(* IEC 61131-3 sources: SortJet_MasterSPS_Aufbau.fbsproj/Device.device.xml.v3^/Plc Logic.plclogic.xml.v3^/Application.application.xml.v3^/09_Station/Shuttle/[151,152] Transfershuttle/0_Konfig, 6 files *)

(* ---- Antriebsinformationen_151.gvl ---- *)
(* METADATA
{
	"v3Meta": {
		"objectGuid": "1be33521-6e58-4da8-829e-a9c5887a7afb"
	}
}
*)
{attribute 'allow_unqualified_access'}
NAMESPACE Antriebsinformationen_151
VAR_GLOBAL

//-------------------------------------------------------------------------------------------------
// ANTRIEBSINFORMATION TRANSFERSHUTTLE
//-------------------------------------------------------------------------------------------------

  apgInfoTransfershuttle151Querfahrt : AntriebsInformationen :=
    (
      wAchsID                                 :=         0,  // Achs ID aus dem EConSet
      stTyp                                   := 'Lateral',  // Typ
      wpSchaltschrank                         :=         2,  // Daten aus dem Schaltplan
      wpSchaltplanreihe                       :=         2,  // Daten aus dem Schaltplan
      wpSchaltplanseite                       :=        60,  // Daten aus dem Schaltplan
      rpMaxGeschwindigkeit                    :=      3333,  // [mm/s]   Max- Geschwindigkeit für den Automatikbetrieb
      rpHandGeschwindigkeit                   :=       200,  // [mm/s]   Hand- Geschwindigkeit
      rpReferenzGeschwindigkeit               :=        50,  // [mm/s]   Geschwindigkeit für die Referenzfahrt
      rpMaxBeschleunigung                     :=      4000,  // [mm/s^2] Max Beschleunigung
      rpMaxVerzoegerung                       :=      4000,  // [mm/s^2] Max Verzoegerung
      rpMaxRuckzeit                           :=       300,  // [ms]     Ruckzeit des Antriebs
      rpReduzierteBeschleunigung              :=      4000,  // [mm/s^2] Reduzierte Beschleunigung
      rpReduzierteVerzoegerung                :=      4000,  // [mm/s^2] Reduzierte Verzoegerung
      rpEinrichtGeschwindigkeit               :=        50,  // [mm/s]   Max Geschwindigkeit während der Einrichtung der Anlage
      rpReduzierteGeschwindigkeit             :=       0.0,  // [mm/s]   Reduzierte Geschwindigkeit
      rpBeschleunigungFremdanlage             :=       0.0,  // [mm/s^2] Beschleunigung zu einer Fremdanlage
      rpGeschwindigkeitMessen                 :=       0.0,  // [mm/s] Geschwindigkeit beim Scheiben messen
      rpGeschwindigkeitSystemcheck            :=     500.0,  // [mm/s]   Geschwindigkeit im Systemcheck (nur Glastransport)
      rpGeschwindigkeitSystemcheckReduzierung :=     167.0,  // [mm/s]   Geschwindigkeit im Systemcheck bei belegtem Vorstop-Sensor (nur Glastransport)
      stOptionen                              := ( eEndschalterQuelle    := Endschalterquelle_EN.UMRICHTER, // Hardware-Endschalter: KEINE, UMRICHTER oder SPS
                                                   bVersorgungUeberXVR   := FALSE,                          // XVR-Modus: brueckt Hauptschalter 400 V und LS 230 V
                                                   bBremseLoesenFreigabe := FALSE )                         // Der Antrieb darf über eine Betriebsart die Bremse lösen
    );

  apgInfoTransfer151Glastransport : ARRAY[cWAND_1..cANZAHL_WAENDE] OF AntriebsInformationen := [
    (
      wAchsID                                 :=         1,  // Achs ID aus dem EConSet
      stTyp                                   :=    'Belt',  // Typ
      wpSchaltschrank                         :=         2,  // Daten aus dem Schaltplan
      wpSchaltplanreihe                       :=         2,  // Daten aus dem Schaltplan
      wpSchaltplanseite                       :=        65,  // Daten aus dem Schaltplan
      rpMaxGeschwindigkeit                    :=       667,  // [mm/s]   Max- Geschwindigkeit für den Automatikbetrieb
      rpHandGeschwindigkeit                   :=       200,  // [mm/s]   Hand- Geschwindigkeit
      rpReduzierteGeschwindigkeit             :=        67,  // [mm/s]   Reduzierte Geschwindigkeit
      rpReferenzGeschwindigkeit               :=         0,  // [mm/s]   Geschwindigkeit für die Referenzfahrt
      rpEinrichtGeschwindigkeit               :=        50,  // [mm/s]   Max Geschwindigkeit während der Einrichtung der Anlage
      rpMaxBeschleunigung                     :=      1500,  // [mm/s^2] Max Beschleunigung
      rpMaxVerzoegerung                       :=      2000,  // [mm/s^2] Max Verzoegerung
      rpMaxRuckzeit                           :=        50,  // [ms]     Ruckzeit des Antriebs
      rpReduzierteBeschleunigung              :=      1000,  // [mm/s^2] Reduzierte Beschleunigung
      rpReduzierteVerzoegerung                :=      1000,  // [mm/s^2] Reduzierte Verzoegerung
      rpBeschleunigungFremdanlage             :=      1000,  // [mm/s^2] Beschleunigung zu einer Fremdanlage
      rpGeschwindigkeitMessen                 :=       667,  // [mm/s] Geschwindigkeit beim Scheiben messen
      rpGeschwindigkeitSystemcheck            :=     500.0,  // [mm/s]   Geschwindigkeit im Systemcheck (nur Glastransport)
      rpGeschwindigkeitSystemcheckReduzierung :=     167.0,  // [mm/s]   Geschwindigkeit im Systemcheck bei belegtem Vorstop-Sensor (nur Glastransport)
      stOptionen                              := ( eEndschalterQuelle    := Endschalterquelle_EN.KEINE,     // Hardware-Endschalter: KEINE, UMRICHTER oder SPS
                                                   bVersorgungUeberXVR   := FALSE,                          // XVR-Modus: brueckt Hauptschalter 400 V und LS 230 V
                                                   bBremseLoesenFreigabe := FALSE )                         // Der Antrieb darf über eine Betriebsart die Bremse lösen
    )];

END_VAR
END_NAMESPACE

(* ---- Antriebsinformationen_152.gvl ---- *)
(* METADATA
{
	"v3Meta": {
		"objectGuid": "34921d73-d8bd-4657-bcb2-03b0c8f4301f"
	}
}
*)
{attribute 'allow_unqualified_access'}
NAMESPACE Antriebsinformationen_152
VAR_GLOBAL

//-------------------------------------------------------------------------------------------------
// ANTRIEBSINFORMATION TRANSFERSHUTTLE
//-------------------------------------------------------------------------------------------------

  apgInfoTransfershuttle152Querfahrt : AntriebsInformationen :=
    (
      wAchsID                                 :=         2,  // Achs ID aus dem EConSet
      stTyp                                   := 'Lateral',  // Typ
      wpSchaltschrank                         :=         2,  // Daten aus dem Schaltplan
      wpSchaltplanreihe                       :=         2,  // Daten aus dem Schaltplan
      wpSchaltplanseite                       :=        60,  // Daten aus dem Schaltplan
      rpMaxGeschwindigkeit                    :=      3333,  // [mm/s]   Max- Geschwindigkeit für den Automatikbetrieb
      rpHandGeschwindigkeit                   :=       200,  // [mm/s]   Hand- Geschwindigkeit
      rpReferenzGeschwindigkeit               :=        50,  // [mm/s]   Geschwindigkeit für die Referenzfahrt
      rpMaxBeschleunigung                     :=      4000,  // [mm/s^2] Max Beschleunigung
      rpMaxVerzoegerung                       :=      4000,  // [mm/s^2] Max Verzoegerung
      rpMaxRuckzeit                           :=       300,  // [ms]     Ruckzeit des Antriebs
      rpReduzierteBeschleunigung              :=      4000,  // [mm/s^2] Reduzierte Beschleunigung
      rpReduzierteVerzoegerung                :=      4000,  // [mm/s^2] Reduzierte Verzoegerung
      rpEinrichtGeschwindigkeit               :=        50,  // [mm/s]   Max Geschwindigkeit während der Einrichtung der Anlage
      rpReduzierteGeschwindigkeit             :=       0.0,  // [mm/s]   Reduzierte Geschwindigkeit
      rpBeschleunigungFremdanlage             :=       0.0,  // [mm/s^2] Beschleunigung zu einer Fremdanlage
      rpGeschwindigkeitMessen                 :=       0.0,  // [mm/s] Geschwindigkeit beim Scheiben messen
      rpGeschwindigkeitSystemcheck            :=     500.0,  // [mm/s]   Geschwindigkeit im Systemcheck (nur Glastransport)
      rpGeschwindigkeitSystemcheckReduzierung :=     167.0,  // [mm/s]   Geschwindigkeit im Systemcheck bei belegtem Vorstop-Sensor (nur Glastransport)
      stOptionen                              := ( eEndschalterQuelle    := Endschalterquelle_EN.UMRICHTER, // Hardware-Endschalter: KEINE, UMRICHTER oder SPS
                                                   bVersorgungUeberXVR   := FALSE,                          // XVR-Modus: brueckt Hauptschalter 400 V und LS 230 V
                                                   bBremseLoesenFreigabe := FALSE )                         // Der Antrieb darf über eine Betriebsart die Bremse lösen
    );

  apgInfoTransfer152Glastransport : ARRAY[cWAND_1..cANZAHL_WAENDE] OF AntriebsInformationen := [
    (
      wAchsID                                 :=         3,  // Achs ID aus dem EConSet
      stTyp                                   :=    'Belt',  // Typ
      wpSchaltschrank                         :=         2,  // Daten aus dem Schaltplan
      wpSchaltplanreihe                       :=         2,  // Daten aus dem Schaltplan
      wpSchaltplanseite                       :=        65,  // Daten aus dem Schaltplan
      rpMaxGeschwindigkeit                    :=       667,  // [mm/s]   Max- Geschwindigkeit für den Automatikbetrieb
      rpHandGeschwindigkeit                   :=       200,  // [mm/s]   Hand- Geschwindigkeit
      rpReduzierteGeschwindigkeit             :=        67,  // [mm/s]   Reduzierte Geschwindigkeit
      rpReferenzGeschwindigkeit               :=         0,  // [mm/s]   Geschwindigkeit für die Referenzfahrt
      rpEinrichtGeschwindigkeit               :=        50,  // [mm/s]   Max Geschwindigkeit während der Einrichtung der Anlage
      rpMaxBeschleunigung                     :=      1500,  // [mm/s^2] Max Beschleunigung
      rpMaxVerzoegerung                       :=      2000,  // [mm/s^2] Max Verzoegerung
      rpMaxRuckzeit                           :=        50,  // [ms]     Ruckzeit des Antriebs
      rpReduzierteBeschleunigung              :=      1000,  // [mm/s^2] Reduzierte Beschleunigung
      rpReduzierteVerzoegerung                :=      1000,  // [mm/s^2] Reduzierte Verzoegerung
      rpBeschleunigungFremdanlage             :=      1000,  // [mm/s^2] Beschleunigung zu einer Fremdanlage
      rpGeschwindigkeitMessen                 :=       667,  // [mm/s] Geschwindigkeit beim Scheiben messen
      rpGeschwindigkeitSystemcheck            :=     500.0,  // [mm/s]   Geschwindigkeit im Systemcheck (nur Glastransport)
      rpGeschwindigkeitSystemcheckReduzierung :=     167.0,  // [mm/s]   Geschwindigkeit im Systemcheck bei belegtem Vorstop-Sensor (nur Glastransport)
      stOptionen                              := ( eEndschalterQuelle    := Endschalterquelle_EN.KEINE,     // Hardware-Endschalter: KEINE, UMRICHTER oder SPS
                                                   bVersorgungUeberXVR   := FALSE,                          // XVR-Modus: brueckt Hauptschalter 400 V und LS 230 V
                                                   bBremseLoesenFreigabe := FALSE )                         // Der Antrieb darf über eine Betriebsart die Bremse lösen
    )];

END_VAR
END_NAMESPACE

(* ---- MK_Transfershuttle_151.gvl ---- *)
(* METADATA
{
	"v3Meta": {
		"objectGuid": "7b0b09af-66f3-4d35-ae87-7c9d4c69f207"
	}
}
*)
{attribute 'allow_unqualified_access'}
NAMESPACE MK_Transfershuttle_151
VAR_GLOBAL

//-------------------------------------------------------------------------------------------------
// TRANSFERSHUTTLE ALLGEMEIN
//-------------------------------------------------------------------------------------------------

  apgMKTransfershuttle151 : Parameter_Station :=
    (
      stStationsNummern                 := ( NummerIntern := 151,                                     // Stationsnummer fuer das MMI und die Stationsangabe der Meldungen
                                             NummerExtern := 1151,                                    // Stationsnummer fuer Bedienermeldungen
                                             NummerSPS    := 151 ),                                   // Stationsnummer SPS-intern (Indizes)
      bDeaktivieren                     := FALSE,                                                     // Station deaktiviert (keine Auftraege, keine Referenzfahrt)
      wMeldungsNummer                   := 350,                                                       // Basis-Meldungsnummer (WatchIO)
      eStationsTyp                      := eTransfershuttle,                                          // Typ der Station
      eaAutomatikkreis                  := [eAutomatikkreis_1, eAutomatikkreis_2],                    // Automatikkreise, zu denen die Station gehoert
      eaSicherheitskreis                := [eSicherheitskreis_1],                                     // Sicherheitskreise, in die die Station eingebunden ist
      // astSicherheitskreisTeilabschaltung
      eSystemcheckZyklus                := eSystemcheckZyklus_1,                                      // In welchem Zyklus des Systemchecks die Station geprueft wird
      stSchnittstellendaten             := ( wVorgaengerStation := cSTATION_DEFAULT,                  // Station vor dieser Station (cSTATION_DYNAMISCH bei mehreren)
                                             wNachfolgerStation := cSTATION_DEFAULT,                  // Station nach dieser Station (cSTATION_DYNAMISCH bei mehreren)
                                             bStationIstShuttle := TRUE ),                            // Station ist ein Shuttle

      stStationsOptionen                := (
                                            stSystemcheck := (
                                              bScheibenVermessenSystemCheck           := FALSE,       // Scheiben im Systemcheck vermessen
                                              bScheibeNachSystemcheckAufAuslauf       := FALSE,       // Scheibe nach dem Systemcheck auf den Auslaufsensor fahren
                                              bSystemCheckMitVorgaengerBatchTransport := FALSE,       // derzeit ohne Funktion
                                              bSystemCheckMitNachfolgerBatchTransport := FALSE,       // derzeit ohne Funktion
                                              bOptionSystemCheckScheibeMittigLegen    := FALSE        // derzeit ohne Funktion
                                            ),

                                            stTransfershuttle := (
                                              bMasterStation                          := TRUE,        // Ob es sich um ein Master (Master-Slave) - Station handelt. Aktuell gebraucht bei Transfershuttle- Verbund
                                              bTransferShuttleFuerFaecherwagen        := FALSE,       // Transfershuttle beschickt Faecherwagen
                                              bTransferShuttleMitUltraschallSensoren  := FALSE,       // Luftabfragen als Ultraschallsensoren (Schliesser)
                                              bTransfershuttleIstVerfahrbarerSpeicher := FALSE        // Transfershuttle ist verfahrbarer Speicher
                                            ),

                                            stGlastransport := (
                                              bVortransport                          := TRUE,         // Vortransport aktivieren [Bsp.: Nach einem Eintransport mit gesetztem Bit <Letzte Scheibe>]
                                              bTransportMasterSlaveEintransport      := FALSE,        // derzeit ohne Funktion
                                              bTransportMasterSlaveAustransport      := TRUE ,        // Austransport als Slave auf die Achse des Nachfolgers
                                              bGLasUebernahmeSenkrecht               := FALSE,        // RKT - Eintransport in Senkrechter-Position bzw. in Waagerechter- Position [default]
                                              bAustransportISOLinie                  := FALSE,        // Austransport an eine ISO-Linie
                                              bScheibenVermessen                     := FALSE,        // Scheibenmessung am Anlegetisch/Anlegewand
                                              bMessrichtungNegativ                   := FALSE,        // Negative Fahrtrichtung beim Messen
                                              bScheibenmessungEintransport           := FALSE,        // Scheibenmessung beim Eintransport
                                              bScheibenmessungSensorVorabAuslauf     := FALSE         // Scheibenmessung mit SensorVorabAuslauf z.B. Anlegewand
                                            ),

                                            // stAnlegetisch
                                            // stEckuebergabe
                                            // stDrehstation
                                            bVorAbKomponentenAnsteuerung            := FALSE,         // VorAbKomponentenAnsteuerung Auftraege werden bearbeitet
                                            bVerstellungEinAusGefahrenLogikDrehen   := FALSE,         // Verstellung: Logik ein-/ausgefahren gedreht
                                            bLangsamfahrtNockenQuerfahrtAktivieren  := FALSE,         // Querfahrt: Langsamfahrt-Nocken auswerten
                                            bSKBlockierenDurchVorabSensoren         := FALSE,         // Vorab-Sensoren belegt blockieren das Oeffnen des Sicherheitskreises
                                            bStationLeerfahrenBeiSkAnforderung      := FALSE,         // Station bei Anforderung Sicherheitskreis leerfahren
                                            bGlasAbgenommenAutomatischQuittieren    := FALSE,         // derzeit ohne Funktion
                                            bScheibeAbnehmenNachEintransport        := FALSE          // Scheibe nach dem Eintransport wieder abnehmen
                                          ),

      stStationsAufbau                  := (
                                            bGeblase                      := [cANZAHL_WAENDE(FALSE)], // Ausbaustufe: Geblaese je Wand
                                            bGlastransport                := [cANZAHL_WAENDE(TRUE)],  // Ausbaustufe: Glastransport je Wand
                                            bKippen                       := [cANZAHL_WAENDE(FALSE)], // Ausbaustufe: Kippen je Wand
                                            bKippenSchuetz                := FALSE,                   // Kippen ueber Schuetz statt Umrichter
                                            bTransportVerstellung         := [cANZAHL_WAENDE(FALSE)], // Ausbaustufe Shuttle: Transport-/Dickenverstellung je Wand
                                            bHub                          := FALSE,                   // Ausbaustufe: Hub der Station
                                            bHubrahmen                    := FALSE,                   // Ausbaustufe: Hubrahmen (Riemen heben/senken)
                                            bDrehen                       := FALSE,                   // Ausbaustufe: Drehen
                                            bQuerachse                    := FALSE,                   // Ausbaustufe: Querachse
                                            bMessachse                    := FALSE,                   // Ausbaustufe: Messachse (Anlegetisch, Anlegewand)
                                            bDruckluft                    := TRUE,                    // Druckluftueberwachung vorhanden
                                            bAnschlag                     := FALSE,                   // Ausbaustufe: Ausrichtanschlaege
                                            bSensorAuslauf                := TRUE,                    // Auslaufsensor vorhanden
                                            bSensorEinlauf                := TRUE,                    // Einlaufsensor vorhanden
                                            bSensorEinlaufStopp           := FALSE,                   // Shuttle: zusaetzlicher Stopp-Sensor am Einlauf (ohne: Einlaufsensor), Gegenstueck zum Auslauf-Stopp im Rueckwaertstransport
                                            bSensorAuslaufStopp           := FALSE,                   // Shuttle: zusaetzlicher Stopp-Sensor am Auslauf (ohne: Auslaufsensor), Verfahrfreigabe und Scheibe hat Shuttle verlassen
                                            bDurchlaufSperreZumNachfolger := FALSE,                   // Ausbaustufe: bewegliche Abschrankung zum Nachfolger
                                            bQuerfahrt                    := TRUE,                    // Ausbaustufe: Querfahrt
                                            bDLSSchmiersystem             := TRUE,                    // Zentralschmierung DLS vorhanden
                                            bWandverstellung              := [ FALSE ],               // Ausbaustufe Station: Wandverstellung je Wand
                                            bWandverstellungMotorisch     := FALSE,                   // Shuttle: Transport-/Wandverstellung mit Antrieb statt pneumatisch
                                            bRoellchenleiste              := [ FALSE ],               // Ausbaustufe Station: Roellchenleiste je Wand
                                            bDurchgang                    := FALSE,                   // Station ist Teil eines Durchgangs (belegt = Oeffnen blockiert)
                                            bSlaveAntrieb                 := FALSE,                   // Glastransport mit Slave-Antrieb
                                            bRolltor                      := FALSE,                   // Ausbaustufe Faecherwagen: Rolltor
                                            bKlemmzylinder                := FALSE,                   // Ausbaustufe Faecherwagen: Klemmzylinder fixiert den Oberrahmen beim Ein- und Ausschleusen
                                            bGreifer                      := [cANZAHL_WAENDE(FALSE)], // Shuttle: Greifer je Wand (Scheibe aus dem Faecherwagen ziehen bzw. hineinschieben)
                                            bRFID                         := FALSE,                   // RFID-Leser vorhanden
                                            bAGV                          := FALSE,                   // Ausbaustufe Faecherwagen: Betrieb mit AGV
                                            bKipparme                     := FALSE,                   // Ausbaustufe: Kipparme
                                            bMessachseAmEndeVomTisch      := FALSE,                   // Messachse am Ende des Tisches (Hoehenfehler fragt den Bediener)
                                            bGlastransportSlaveVorhanden  := FALSE,                   // Glastransport mit Slave-Antrieb (Meldungen/Ueberwachung Slave)
                                            wHydraulikstation             := 0                        // Faecherwagen Hydraulik: zugeordnete Hydraulikstation (cHYDRAULIKSTATION_x), 0 = keine
                                          ),

      stStationsParameter               := (
                                            rLaengeUebergroesseScheibe              := 4240,          // Shuttle: ab dieser Scheibenlaenge gilt die Scheibe als uebergross [mm]
                                            rMinGlasHoeheAutomatischenEintransport  := 500,           // VSG: Mindesthoehe fuer automatischen Eintransport [mm]
                                            rMinGlasLaengeAutomatischenEintransport := 500,           // VSG: Mindestlaenge fuer automatischen Eintransport [mm]
                                            wMaximaleAnzahlAktiverAuftraege         := 1,             // derzeit ohne Funktion
                                            rMinPosSwEsEingrenzung                  := 0.0,           // Externer zusaetzlicher Software-Endschalter MIN; 0 = inaktiv; darf den MK-MIN nur weiter eingrenzen
                                            rMaxPosSwEsEingrenzung                  := 0.0,           // Externer zusaetzlicher Software-Endschalter MAX; 0 = inaktiv; darf den MK-MAX nur weiter eingrenzen
                                            rPosFreigabePufferAusfahren             := 0.0            // derzeit ohne Funktion
                                          ),

      // stFremdanlage
      stGlasdaten                       := [
                                            (
                                              rlMinGlasLaenge := 350,                                 // minimal zulässige GlasLänge
                                              rlMaxGlasLaenge := 2500,                                // maximale zulässige GlasLänge
                                              rlMinGlasHoehe  := 190,                                 // minimal zulässige GlasHöhe
                                              rlMaxGlasHoehe  := 1800,                                // maximale zulässige GlasHöhe
                                              rlMinGlasDicke  := 3,                                 // minimal zulässige GlasDicke
                                              rlMaxGlasDicke  := 12.76,                                  // maximal zulaessige Glasdicke [mm]
                                              rlLaengeMaxGlas := 0.0                                  // maximal zulaessige Glaslaenge [mm]
                                            )]
      // astShuttleAnhaltenQuellen
    );

//-------------------------------------------------------------------------------------------------
// TRANSFERSHUTTLE GLASTRANSPORT
//-------------------------------------------------------------------------------------------------

  apgTransfer151Glastransport : ARRAY[cWAND_1..cANZAHL_WAENDE] OF Parameter_TransfershuttleGlastransport := [
    (
      rlLaengeStation                    := 3945, // Länge der Station
      rStopFreiFahren                    := 300,  // So weit soll die Scheibe beim Austransport länger fahren
      rWegUeberEinlaufEintransport       := 170,  // Eintransport vorwaerts: Abstand Scheibenhinterkante zum Einlaufsensor [mm]
      rWegUeberEinlaufAustransport       := 50,   // Lage Auf Einlauf: Scheibe liegt um diesen Weg auf dem Einlaufsensor [mm]
      rWegUeberAuslaufEintransport       := 50,   // Eintransport rueckwaerts: Abstand Scheibenhinterkante zum Auslaufsensor [mm]
      rWegUeberAuslaufAustransport       := 50,   // Lage Auf Auslauf: Weg ueber den Auslaufsensor hinaus [mm]
      wEnergieSparZeit                   := 180,  // in Sec, Zeitspanne nach der, der Antrieb deaktiviert wird wenn er keinen Auftrag hat
      rMaxPosAuslaufSensorFreiFahren     := 300,  // Bestimmt die Strecke die Maximal zurueck gefahren werden soll bis der Auslaufsensor  wieder frei ist
      rMaxPosEinlaufSensorFreiFahren     := 300,  // So weit darf maximal der Einlaufsensor frei gefahren weirden
      rgAbstandLuftAbfrageAuslaufShuttle := 0     // Abstand in mm von der Einlaufluftschranke zum Inputshuttle Auslaufsensor
    )];

END_VAR
END_NAMESPACE

(* ---- MK_Transfershuttle_152.gvl ---- *)
(* METADATA
{
	"v3Meta": {
		"objectGuid": "e51deda7-4c76-464f-a8c8-8f73f5e7edb3"
	}
}
*)
{attribute 'allow_unqualified_access'}
NAMESPACE MK_Transfershuttle_152
VAR_GLOBAL

//-------------------------------------------------------------------------------------------------
// TRANSFERSHUTTLE ALLGEMEIN
//-------------------------------------------------------------------------------------------------

  apgMKTransfershuttle152 : Parameter_Station :=
    (
      stStationsNummern                 := ( NummerIntern := 152,                                     // Stationsnummer fuer das MMI und die Stationsangabe der Meldungen
                                             NummerExtern := 1152,                                    // Stationsnummer fuer Bedienermeldungen
                                             NummerSPS    := 152 ),                                   // Stationsnummer SPS-intern (Indizes)
      bDeaktivieren                     := FALSE,                                                     // Station deaktiviert (keine Auftraege, keine Referenzfahrt)
      wMeldungsNummer                   := 380,                                                       // Basis-Meldungsnummer (WatchIO)
      eStationsTyp                      := eTransfershuttle,                                          // Typ der Station
      eaAutomatikkreis                  := [eAutomatikkreis_1, eAutomatikkreis_2],                    // Automatikkreise, zu denen die Station gehoert
      eaSicherheitskreis                := [eSicherheitskreis_1],                                     // Sicherheitskreise, in die die Station eingebunden ist
      // astSicherheitskreisTeilabschaltung
      eSystemcheckZyklus                := eSystemcheckZyklus_1,                                      // In welchem Zyklus des Systemchecks die Station geprueft wird
      stSchnittstellendaten             := ( wVorgaengerStation := cSTATION_DEFAULT,                  // Station vor dieser Station (cSTATION_DYNAMISCH bei mehreren)
                                             wNachfolgerStation := cSTATION_DEFAULT,                  // Station nach dieser Station (cSTATION_DYNAMISCH bei mehreren)
                                             bStationIstShuttle := TRUE ),                            // Station ist ein Shuttle

      stStationsOptionen                := (
                                            stSystemcheck := (
                                              bScheibenVermessenSystemCheck           := FALSE,       // Scheiben im Systemcheck vermessen
                                              bScheibeNachSystemcheckAufAuslauf       := FALSE,       // Scheibe nach dem Systemcheck auf den Auslaufsensor fahren
                                              bSystemCheckMitVorgaengerBatchTransport := FALSE,       // derzeit ohne Funktion
                                              bSystemCheckMitNachfolgerBatchTransport := FALSE,       // derzeit ohne Funktion
                                              bOptionSystemCheckScheibeMittigLegen    := FALSE        // derzeit ohne Funktion
                                            ),

                                            stTransfershuttle := (
                                              bMasterStation                          := TRUE,        // Ob es sich um ein Master (Master-Slave) - Station handelt. Aktuell gebraucht bei Transfershuttle- Verbund
                                              bTransferShuttleFuerFaecherwagen        := FALSE,       // Transfershuttle beschickt Faecherwagen
                                              bTransferShuttleMitUltraschallSensoren  := FALSE,       // Luftabfragen als Ultraschallsensoren (Schliesser)
                                              bTransfershuttleIstVerfahrbarerSpeicher := FALSE        // Transfershuttle ist verfahrbarer Speicher
                                            ),

                                            stGlastransport := (
                                              bVortransport                          := TRUE,         // Vortransport aktivieren [Bsp.: Nach einem Eintransport mit gesetztem Bit <Letzte Scheibe>]
                                              bTransportMasterSlaveEintransport      := FALSE,        // derzeit ohne Funktion
                                              bTransportMasterSlaveAustransport      := TRUE ,        // Austransport als Slave auf die Achse des Nachfolgers
                                              bGLasUebernahmeSenkrecht               := FALSE,        // RKT - Eintransport in Senkrechter-Position bzw. in Waagerechter- Position [default]
                                              bAustransportISOLinie                  := FALSE,        // Austransport an eine ISO-Linie
                                              bScheibenVermessen                     := FALSE,        // Scheibenmessung am Anlegetisch/Anlegewand
                                              bMessrichtungNegativ                   := FALSE,        // Negative Fahrtrichtung beim Messen
                                              bScheibenmessungEintransport           := FALSE,        // Scheibenmessung beim Eintransport
                                              bScheibenmessungSensorVorabAuslauf     := FALSE         // Scheibenmessung mit SensorVorabAuslauf z.B. Anlegewand
                                            ),

                                            // stAnlegetisch
                                            // stEckuebergabe
                                            // stDrehstation
                                            bVorAbKomponentenAnsteuerung            := FALSE,         // VorAbKomponentenAnsteuerung Auftraege werden bearbeitet
                                            bVerstellungEinAusGefahrenLogikDrehen   := FALSE,         // Verstellung: Logik ein-/ausgefahren gedreht
                                            bLangsamfahrtNockenQuerfahrtAktivieren  := FALSE,         // Querfahrt: Langsamfahrt-Nocken auswerten
                                            bSKBlockierenDurchVorabSensoren         := FALSE,         // Vorab-Sensoren belegt blockieren das Oeffnen des Sicherheitskreises
                                            bStationLeerfahrenBeiSkAnforderung      := FALSE,         // Station bei Anforderung Sicherheitskreis leerfahren
                                            bGlasAbgenommenAutomatischQuittieren    := FALSE,         // derzeit ohne Funktion
                                            bScheibeAbnehmenNachEintransport        := FALSE          // Scheibe nach dem Eintransport wieder abnehmen
                                          ),

      stStationsAufbau                  := (
                                            bGeblase                      := [cANZAHL_WAENDE(FALSE)], // Ausbaustufe: Geblaese je Wand
                                            bGlastransport                := [cANZAHL_WAENDE(TRUE)],  // Ausbaustufe: Glastransport je Wand
                                            bKippen                       := [cANZAHL_WAENDE(FALSE)], // Ausbaustufe: Kippen je Wand
                                            bKippenSchuetz                := FALSE,                   // Kippen ueber Schuetz statt Umrichter
                                            bTransportVerstellung         := [cANZAHL_WAENDE(FALSE)], // Ausbaustufe Shuttle: Transport-/Dickenverstellung je Wand
                                            bHub                          := FALSE,                   // Ausbaustufe: Hub der Station
                                            bHubrahmen                    := FALSE,                   // Ausbaustufe: Hubrahmen (Riemen heben/senken)
                                            bDrehen                       := FALSE,                   // Ausbaustufe: Drehen
                                            bQuerachse                    := FALSE,                   // Ausbaustufe: Querachse
                                            bMessachse                    := FALSE,                   // Ausbaustufe: Messachse (Anlegetisch, Anlegewand)
                                            bDruckluft                    := TRUE,                    // Druckluftueberwachung vorhanden
                                            bAnschlag                     := FALSE,                   // Ausbaustufe: Ausrichtanschlaege
                                            bSensorAuslauf                := TRUE,                    // Auslaufsensor vorhanden
                                            bSensorEinlauf                := TRUE,                    // Einlaufsensor vorhanden
                                            bSensorEinlaufStopp           := FALSE,                   // Shuttle: zusaetzlicher Stopp-Sensor am Einlauf (ohne: Einlaufsensor), Gegenstueck zum Auslauf-Stopp im Rueckwaertstransport
                                            bSensorAuslaufStopp           := FALSE,                   // Shuttle: zusaetzlicher Stopp-Sensor am Auslauf (ohne: Auslaufsensor), Verfahrfreigabe und Scheibe hat Shuttle verlassen
                                            bDurchlaufSperreZumNachfolger := FALSE,                   // Ausbaustufe: bewegliche Abschrankung zum Nachfolger
                                            bQuerfahrt                    := TRUE,                    // Ausbaustufe: Querfahrt
                                            bDLSSchmiersystem             := TRUE,                    // Zentralschmierung DLS vorhanden
                                            bWandverstellung              := [ FALSE ],               // Ausbaustufe Station: Wandverstellung je Wand
                                            bWandverstellungMotorisch     := FALSE,                   // Shuttle: Transport-/Wandverstellung mit Antrieb statt pneumatisch
                                            bRoellchenleiste              := [ FALSE ],               // Ausbaustufe Station: Roellchenleiste je Wand
                                            bDurchgang                    := FALSE,                   // Station ist Teil eines Durchgangs (belegt = Oeffnen blockiert)
                                            bSlaveAntrieb                 := FALSE,                   // Glastransport mit Slave-Antrieb
                                            bRolltor                      := FALSE,                   // Ausbaustufe Faecherwagen: Rolltor
                                            bKlemmzylinder                := FALSE,                   // Ausbaustufe Faecherwagen: Klemmzylinder fixiert den Oberrahmen beim Ein- und Ausschleusen
                                            bGreifer                      := [cANZAHL_WAENDE(FALSE)], // Shuttle: Greifer je Wand (Scheibe aus dem Faecherwagen ziehen bzw. hineinschieben)
                                            bRFID                         := FALSE,                   // RFID-Leser vorhanden
                                            bAGV                          := FALSE,                   // Ausbaustufe Faecherwagen: Betrieb mit AGV
                                            bKipparme                     := FALSE,                   // Ausbaustufe: Kipparme
                                            bMessachseAmEndeVomTisch      := FALSE,                   // Messachse am Ende des Tisches (Hoehenfehler fragt den Bediener)
                                            bGlastransportSlaveVorhanden  := FALSE,                   // Glastransport mit Slave-Antrieb (Meldungen/Ueberwachung Slave)
                                            wHydraulikstation             := 0                        // Faecherwagen Hydraulik: zugeordnete Hydraulikstation (cHYDRAULIKSTATION_x), 0 = keine
                                          ),

      stStationsParameter               := (
                                            rLaengeUebergroesseScheibe              := 4240,          // Shuttle: ab dieser Scheibenlaenge gilt die Scheibe als uebergross [mm]
                                            rMinGlasHoeheAutomatischenEintransport  := 500,           // VSG: Mindesthoehe fuer automatischen Eintransport [mm]
                                            rMinGlasLaengeAutomatischenEintransport := 500,           // VSG: Mindestlaenge fuer automatischen Eintransport [mm]
                                            wMaximaleAnzahlAktiverAuftraege         := 1,             // derzeit ohne Funktion
                                            rMinPosSwEsEingrenzung                  := 0.0,           // Externer zusaetzlicher Software-Endschalter MIN; 0 = inaktiv; darf den MK-MIN nur weiter eingrenzen
                                            rMaxPosSwEsEingrenzung                  := 0.0,           // Externer zusaetzlicher Software-Endschalter MAX; 0 = inaktiv; darf den MK-MAX nur weiter eingrenzen
                                            rPosFreigabePufferAusfahren             := 0.0            // derzeit ohne Funktion
                                          ),

      // stFremdanlage
      stGlasdaten                       := [
                                            (
                                              rlMinGlasLaenge := 350,                                 // minimal zulässige GlasLänge
                                              rlMaxGlasLaenge := 2500,                                // maximale zulässige GlasLänge
                                              rlMinGlasHoehe  := 190,                                 // minimal zulässige GlasHöhe
                                              rlMaxGlasHoehe  := 1800,                                // maximale zulässige GlasHöhe
                                              rlMinGlasDicke  := 3,                                 // minimal zulässige GlasDicke
                                              rlMaxGlasDicke  := 12.76,                                  // maximal zulaessige Glasdicke [mm]
                                              rlLaengeMaxGlas := 0.0                                  // maximal zulaessige Glaslaenge [mm]
                                            )]
      // astShuttleAnhaltenQuellen
    );

//-------------------------------------------------------------------------------------------------
// TRANSFERSHUTTLE GLASTRANSPORT
//-------------------------------------------------------------------------------------------------

  apgTransfer152Glastransport : ARRAY[cWAND_1..cANZAHL_WAENDE] OF Parameter_TransfershuttleGlastransport := [
    (
      rlLaengeStation                    := 3945, // Länge der Station
      rStopFreiFahren                    := 300,  // So weit soll die Scheibe beim Austransport länger fahren
      rWegUeberEinlaufEintransport       := 170,   // Eintransport vorwaerts: Abstand Scheibenhinterkante zum Einlaufsensor [mm]
      rWegUeberEinlaufAustransport       := 50,   // Lage Auf Einlauf: Scheibe liegt um diesen Weg auf dem Einlaufsensor [mm]
      rWegUeberAuslaufEintransport       := 50,   // Eintransport rueckwaerts: Abstand Scheibenhinterkante zum Auslaufsensor [mm]
      rWegUeberAuslaufAustransport       := 50,   // Lage Auf Auslauf: Weg ueber den Auslaufsensor hinaus [mm]
      wEnergieSparZeit                   := 180,  // in Sec, Zeitspanne nach der, der Antrieb deaktiviert wird wenn er keinen Auftrag hat
      rMaxPosAuslaufSensorFreiFahren     := 300,  // Bestimmt die Strecke die Maximal zurueck gefahren werden soll bis der Auslaufsensor  wieder frei ist
      rMaxPosEinlaufSensorFreiFahren     := 300,  // So weit darf maximal der Einlaufsensor frei gefahren weirden
      rgAbstandLuftAbfrageAuslaufShuttle := 0     // Abstand in mm von der Einlaufluftschranke zum Inputshuttle Auslaufsensor
    )];

END_VAR
END_NAMESPACE

(* ---- Konfiguration_151.gvl ---- *)
(* METADATA
{
	"v3Meta": {
		"objectGuid": "72743bf1-0a30-469b-b165-3b7b28535a8f"
	}
}
*)
{attribute 'allow_unqualified_access'}
NAMESPACE Konfiguration_151
VAR_CONFIG
//-------------------------------------------------------------------------------------------------
// KONFIGURATION: BAUSTEIN IO´s
//-------------------------------------------------------------------------------------------------

  // Leitungsschutzschalter
  Globale_Bausteine.aTransfershuttles[151].in_bLeitungsschutz_Querfahrt_OK                                     AT %IX0.7    : BOOL; // IO-L - 151 Querfahrt Sicherung
  Globale_Bausteine.aTransfershuttles[151].in_bDruckluftWartungseinheitOK                                      AT %IX3.1    : BOOL; // IO-L - 151 - 152 Druckluft OK

END_VAR

END_NAMESPACE

(* ---- Konfiguration_152.gvl ---- *)
(* METADATA
{
	"v3Meta": {
		"objectGuid": "67cd098f-c677-47e0-bd7e-f7cb39be9438"
	}
}
*)
{attribute 'allow_unqualified_access'}
NAMESPACE Konfiguration_152
VAR_CONFIG
//-------------------------------------------------------------------------------------------------
// KONFIGURATION: BAUSTEIN IO´s
//-------------------------------------------------------------------------------------------------

  // Leitungsschutzschalter
  Globale_Bausteine.aTransfershuttles[152].in_bLeitungsschutz_Querfahrt_OK                                     AT %IX1.0    : BOOL; // IO-L - 152 Querfahrt Sicherung
  Globale_Bausteine.aTransfershuttles[152].in_bDruckluftWartungseinheitOK                                      AT %IX3.1    : BOOL; // IO-L - 151 - 152 Druckluft OK

END_VAR

END_NAMESPACE
